(* IEC 61131-3 sources: packers-hmi/plc, 2 files *)

(* ---- ST_Analog.st ---- *)
// Analog value with range and engineering units, modeled on OPC UA's AnalogItem.
// Used for both setpoints and process values:
//   Setpoint:      fMin/fMax = allowed entry range. The HMI rejects out-of-range entries, the PLC enforces it.
//   Process value: fMin/fMax = instrument range (for bar graphs, gauges, trend scaling).
// Whether the HMI can write it comes from {attribute 'hmi_write'}, not from this type.
// On a writable instance, the HMI may write fValue only. fMin, fMax and sEU stay PLC-owned.
TYPE ST_Analog :
STRUCT
    fValue : REAL;
    fMin   : REAL;
    fMax   : REAL;
    sEU    : WSTRING(15);   // Engineering units. WSTRING so °F, µS/cm, m³/h display correctly.
END_STRUCT
END_TYPE

(* ---- GVL_HMI.st ---- *)
// Everything the HMI can see. The server reads this list from the PLC at startup
// and again after every download or online change, so there is no tag list to maintain elsewhere.
//
// {attribute 'hmi_write'} on the line above a variable makes it writable from the HMI.
//   Plain variable (BOOL, REAL, ...): the HMI writes the variable itself.
//   ST_Analog:                        the HMI writes fValue only.
{attribute 'qualified_only'}
VAR_GLOBAL
    // --- Commands: HMI sets TRUE, PLC acts and clears ---
    {attribute 'hmi_write'}
    bStartCmd   : BOOL;
    {attribute 'hmi_write'}
    bStopCmd    : BOOL;

    // --- Status ---
    bRunning    : BOOL;
    nBatchCount : DINT;

    // --- Analog values ---
    {attribute 'hmi_write'}
    stSpeedSP   : ST_Analog := (fValue := 250, fMin := 0, fMax := 500, sEU := "ft/min");   // operator setpoint
    stSpeedPV   : ST_Analog := (fMin := 0, fMax := 600, sEU := "ft/min");                   // measured speed
END_VAR

// =====================================================================
// In MAIN (or the relevant program)
// =====================================================================

// Momentary commands. Stop wins if both arrive in the same scan.
IF GVL_HMI.bStopCmd THEN
    GVL_HMI.bRunning := FALSE;
    GVL_HMI.bStopCmd := FALSE;
ELSIF GVL_HMI.bStartCmd THEN
    GVL_HMI.bRunning := TRUE;
    GVL_HMI.bStartCmd := FALSE;
END_IF

// Enforce setpoint limits in the PLC. The HMI's range check is only a convenience for the operator.
GVL_HMI.stSpeedSP.fValue := LIMIT(GVL_HMI.stSpeedSP.fMin, GVL_HMI.stSpeedSP.fValue, GVL_HMI.stSpeedSP.fMax);
